Staubli VAL3: HMI_action.dtx

mdesc mNomSpeed
string sActionList
public string sIOList
string sSelList
string sSelIO[6]
public string sComment
bool bBack
bool bConfirm
num nSelList
string sLastList
bool bOnsave
public actItem aEditItem
  [0]
    string sComment
    actionItem aActItem[6]
      [0]
        num nIOindex
        num nboolValue
        num nPulseValue
        string sIOtype
        string sValue
        bool bActive
      [1]
        num nIOindex
        num nboolValue
        num nPulseValue
        string sIOtype
        string sValue
        bool bActive
      [2]
        num nIOindex
        num nboolValue
        num nPulseValue
        string sIOtype
        string sValue
        bool bActive
      [3]
        num nIOindex
        num nboolValue
        num nPulseValue
        string sIOtype
        string sValue
        bool bActive
      [4]
        num nIOindex
        num nboolValue
        num nPulseValue
        string sIOtype
        string sValue
        bool bActive
      [5]
        num nIOindex
        num nboolValue
        num nPulseValue
        string sIOtype
        string sValue
        bool bActive
